Fanuc KAREL source: KT00822.KL

PROGRAM KT00822
%NOLOCKGROUP
VAR
  R1: REAL
  R2: REAL
  OUT: INTEGER
BEGIN
  R1 = 2.0
  R2 = 3.0
  R1 = 2.0
  R2 = 3.0
  OUT = SIN(R1)
END KT00822
